FUNCTION_BLOCK Gerador_Generico_HMI (* Service Interface Function Block Type *)
  (* Standard: 61499-2 *)
  (* Version 1.1, 15/10/2026, Hidryco, Hidryco, IHM do Gerador_Generico *)
  PACKAGE Hidryco.HidrycoLib;
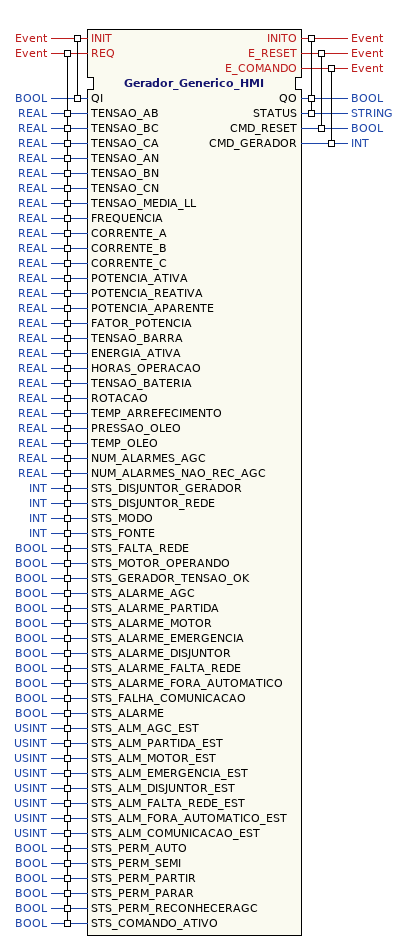
  EVENT_INPUT
    INIT WITH QI;
    REQ WITH TENSAO_AB, TENSAO_BC, TENSAO_CA, TENSAO_AN, TENSAO_BN, TENSAO_CN, TENSAO_MEDIA_LL, FREQUENCIA, CORRENTE_A, CORRENTE_B, CORRENTE_C, POTENCIA_ATIVA, POTENCIA_REATIVA, POTENCIA_APARENTE, FATOR_POTENCIA, TENSAO_BARRA, ENERGIA_ATIVA, HORAS_OPERACAO, TENSAO_BATERIA, ROTACAO, TEMP_ARREFECIMENTO, PRESSAO_OLEO, TEMP_OLEO, NUM_ALARMES_AGC, NUM_ALARMES_NAO_REC_AGC, STS_DISJUNTOR_GERADOR, STS_DISJUNTOR_REDE, STS_MODO, STS_FONTE, STS_FALTA_REDE, STS_MOTOR_OPERANDO, STS_GERADOR_TENSAO_OK, STS_ALARME_AGC, STS_ALARME_PARTIDA, STS_ALARME_MOTOR, STS_ALARME_EMERGENCIA, STS_ALARME_DISJUNTOR, STS_ALARME_FALTA_REDE, STS_ALARME_FORA_AUTOMATICO, STS_FALHA_COMUNICACAO, STS_ALARME, STS_ALM_AGC_EST, STS_ALM_PARTIDA_EST, STS_ALM_MOTOR_EST, STS_ALM_EMERGENCIA_EST, STS_ALM_DISJUNTOR_EST, STS_ALM_FALTA_REDE_EST, STS_ALM_FORA_AUTOMATICO_EST, STS_ALM_COMUNICACAO_EST, STS_PERM_AUTO, STS_PERM_SEMI, STS_PERM_PARTIR, STS_PERM_PARAR, STS_PERM_RECONHECERAGC, STS_COMANDO_ATIVO; (* Atualizacao de status *)
  END_EVENT
  EVENT_OUTPUT
    INITO WITH QO, STATUS;
    E_RESET WITH CMD_RESET;
    E_COMANDO WITH CMD_GERADOR;
  END_EVENT
  VAR_INPUT
    QI : BOOL;
    TENSAO_AB : REAL; (* Tensao A-B (V) *)
    TENSAO_BC : REAL; (* Tensao B-C (V) *)
    TENSAO_CA : REAL; (* Tensao C-A (V) *)
    TENSAO_AN : REAL; (* Tensao A-N (V) *)
    TENSAO_BN : REAL; (* Tensao B-N (V) *)
    TENSAO_CN : REAL; (* Tensao C-N (V) *)
    TENSAO_MEDIA_LL : REAL; (* Tensao media fase-fase (V) *)
    FREQUENCIA : REAL; (* Frequencia (Hz) *)
    CORRENTE_A : REAL; (* Corrente fase A (A) *)
    CORRENTE_B : REAL; (* Corrente fase B (A) *)
    CORRENTE_C : REAL; (* Corrente fase C (A) *)
    POTENCIA_ATIVA : REAL; (* Potencia ativa (kW) *)
    POTENCIA_REATIVA : REAL; (* Potencia reativa (kVAr) *)
    POTENCIA_APARENTE : REAL; (* Potencia aparente (kVA) *)
    FATOR_POTENCIA : REAL; (* Fator de potencia *)
    TENSAO_BARRA : REAL; (* Tensao do lado B (barramento/rede) L1-L2 (V) *)
    ENERGIA_ATIVA : REAL; (* Energia ativa exportada (kWh) *)
    HORAS_OPERACAO : REAL; (* Horas de funcionamento (h) *)
    TENSAO_BATERIA : REAL; (* Tensao da bateria (V) *)
    ROTACAO : REAL; (* Rotacao do motor (rpm) *)
    TEMP_ARREFECIMENTO : REAL; (* Temperatura do liquido de arrefecimento (°C) *)
    PRESSAO_OLEO : REAL; (* Pressao do oleo (bar) *)
    TEMP_OLEO : REAL; (* Temperatura do oleo (°C) *)
    NUM_ALARMES_AGC : REAL; (* Alarmes ativos no AGC *)
    NUM_ALARMES_NAO_REC_AGC : REAL; (* Alarmes nao reconhecidos no AGC *)
    STS_DISJUNTOR_GERADOR : INT; (* Disjuntor do gerador (GB): 0 indefinido/sem comunicacao, 1 aberto, 2 fechado *)
    STS_DISJUNTOR_REDE : INT; (* Disjuntor de rede (MB): 0 indefinido/sem comunicacao, 1 aberto, 2 fechado *)
    STS_MODO : INT; (* Modo do AGC: 0 indefinido, 1 automatico, 2 semi-automatico, 3 manual, 4 bloqueio, 5 teste *)
    STS_FONTE : INT; (* Fonte da saida do QTA: 0 sem fonte, 1 rede, 2 gerador, 3 indefinida (sem comunicacao) *)
    STS_FALTA_REDE : BOOL; (* Falta de rede (AMF) *)
    STS_MOTOR_OPERANDO : BOOL; (* Motor em operacao *)
    STS_GERADOR_TENSAO_OK : BOOL; (* Tensao e frequencia do gerador OK *)
    STS_ALARME_AGC : BOOL; (* Alarme ativo no controlador do gerador (AGC 150) *)
    STS_ALARME_PARTIDA : BOOL; (* Falha na partida do gerador *)
    STS_ALARME_MOTOR : BOOL; (* Desligamento do motor (ECU ou sobrevelocidade) *)
    STS_ALARME_EMERGENCIA : BOOL; (* Parada de emergência do gerador acionada *)
    STS_ALARME_DISJUNTOR : BOOL; (* Falha de disjuntor no QTA (gerador ou rede) *)
    STS_ALARME_FALTA_REDE : BOOL; (* Falta de rede no QTA *)
    STS_ALARME_FORA_AUTOMATICO : BOOL; (* Gerador fora do modo automático *)
    STS_FALHA_COMUNICACAO : BOOL; (* Falha de comunicacao *)
    STS_ALARME : BOOL; (* Algum alarme do gerador *)
    STS_ALM_AGC_EST : USINT; (* Estado do ALARM_BIT Alarme ativo no controlador do gerador (AGC 150) (0 normal, 1 ativo reconhecido, 2 ativo nao reconhecido, 3 saiu nao reconhecido, 4 ativo e saiu nao reconhecido) *)
    STS_ALM_PARTIDA_EST : USINT; (* Estado do ALARM_BIT Falha na partida do gerador (0 normal, 1 ativo reconhecido, 2 ativo nao reconhecido, 3 saiu nao reconhecido, 4 ativo e saiu nao reconhecido) *)
    STS_ALM_MOTOR_EST : USINT; (* Estado do ALARM_BIT Desligamento do motor (ECU ou sobrevelocidade) (0 normal, 1 ativo reconhecido, 2 ativo nao reconhecido, 3 saiu nao reconhecido, 4 ativo e saiu nao reconhecido) *)
    STS_ALM_EMERGENCIA_EST : USINT; (* Estado do ALARM_BIT Parada de emergência do gerador acionada (0 normal, 1 ativo reconhecido, 2 ativo nao reconhecido, 3 saiu nao reconhecido, 4 ativo e saiu nao reconhecido) *)
    STS_ALM_DISJUNTOR_EST : USINT; (* Estado do ALARM_BIT Falha de disjuntor no QTA (gerador ou rede) (0 normal, 1 ativo reconhecido, 2 ativo nao reconhecido, 3 saiu nao reconhecido, 4 ativo e saiu nao reconhecido) *)
    STS_ALM_FALTA_REDE_EST : USINT; (* Estado do ALARM_BIT Falta de rede no QTA (0 normal, 1 ativo reconhecido, 2 ativo nao reconhecido, 3 saiu nao reconhecido, 4 ativo e saiu nao reconhecido) *)
    STS_ALM_FORA_AUTOMATICO_EST : USINT; (* Estado do ALARM_BIT Gerador fora do modo automático (0 normal, 1 ativo reconhecido, 2 ativo nao reconhecido, 3 saiu nao reconhecido, 4 ativo e saiu nao reconhecido) *)
    STS_ALM_COMUNICACAO_EST : USINT; (* Estado do ALARM_BIT falha de comunicacao (0 normal, 1 ativo reconhecido, 2 ativo nao reconhecido, 3 saiu nao reconhecido, 4 ativo e saiu nao reconhecido) *)
    STS_PERM_AUTO : BOOL; (* Comando Auto permitido *)
    STS_PERM_SEMI : BOOL; (* Comando Semi permitido *)
    STS_PERM_PARTIR : BOOL; (* Comando Partir permitido *)
    STS_PERM_PARAR : BOOL; (* Comando Parar permitido *)
    STS_PERM_RECONHECERAGC : BOOL; (* Comando ReconhecerAGC permitido *)
    STS_COMANDO_ATIVO : BOOL; (* Comando sendo enviado ao AGC *)
  END_VAR
  VAR_OUTPUT
    QO : BOOL; (* Event Output Qualifier *)
    STATUS : STRING; (* Service Status *)
    CMD_RESET : BOOL; (* Reconhece os alarmes do gerador *)
    CMD_GERADOR : INT; (* Comando para o AGC: 1 automatico, 2 semiautomatico, 3 partir, 4 parar, 5 reconhecer alarmes do AGC *)
  END_VAR
  SERVICE /
    SEQUENCE 
    END_SEQUENCE
  END_SERVICE
END_FUNCTION_BLOCK
